// TIA Portal V19 export
TYPE "ST_Bit"
   STRUCT
      Bit_0 : Bool;
      Bit_1 : Bool;
      Bit_2 : Bool;
      Bit_3 : Bool;
      Bit_4 : Bool;
      Bit_5 : Bool;
      Bit_6 : Bool;
      Bit_7 : Bool;
   END_STRUCT;
END_TYPE
